(*
See the Beckhoff homepage_ for more information.

Please contact the `Beckhoff Support`_ for technical assistance.

.. _homepage: http://www.beckhoff.de
.. _Beckhoff Support: support@beckhoff.com

For more information see the `PLC Lib Tc2_System`_ and `PLC Lib Tc2_Standard`_.

.. _PLC Lib Tc2_System: https://download.beckhoff.com/download/document/automation/twincat3/TwinCAT_3_PLC_Lib_Tc2_System_EN.pdf
.. _PLC Lib Tc2_Standard: https://download.beckhoff.com/download/document/automation/twincat3/TwinCAT_3_PLC_Lib__Tc2_Standard_EN.pdf

External hyperlinks, like `Beckhoff <http://www.beckhoff.de/>`_.


**Standalone hyperlinks**

See http://www.beckhoff.de for info.

Contact support@beckhoff.com


**Embedded URIs and aliases**

See the `Beckhoff homepage <http://www.beckhoff.de>`_ for info.

This `link <Beckhoff homepage_>`_ is an alias to the link above.


See the `Beckhoff homepage`_ for info.

This link_ is an alias to the link above.

.. _Beckhoff homepage: http://www.beckhoff.de
.. _link: `Beckhoff homepage`_

*)

FUNCTION_BLOCK FB_Libdoc_ExternalHyperlinks
VAR_INPUT
    nVarA : INT;
    nVarB : INT;
END_VAR
VAR_OUTPUT
    nSum : INT;
END_VAR
VAR
END_VAR

END_FUNCTION_BLOCK

(* stored: Version 1.1.0.1, ProductVersion 3.1.4024.0
   POU FB_Libdoc_ExternalHyperlinks: Id {af1f6adf-277a-483c-bc55-8755a439ade6}, SpecialFunc None *)
